(* IEC 61131-3 sources: horner-cscape-mcp/artifacts/projects/Fail_Ladder_Location_Proj/pous, 1 file *)

(* ---- POU_LadderInjection.st ---- *)
PROGRAM POU_LadderInjection
VAR
    InSensor : BOOL := FALSE;
    OutMotor : BOOL;
END_VAR

---[ ]--- InSensor
END_PROGRAM
